// TIA Portal V20 export
// export: Created 2026-10-12T05:35:25.4874233Z, ExportSetting WithDefaults, DisplayName Totally Integrated Automation Portal, DisplayVersion V20, DisplayName TIA Portal Openness, DisplayVersion V20, DisplayName TIA Portal Teamcenter Gateway, DisplayVersion V20, DisplayName TIA Portal Version Control Interface, DisplayVersion V20, DisplayName SINAMICS Startdrive Advanced, DisplayVersion V20 SP1 Update 2, DisplayName SINAMICS Startdrive G110M, G120, G120C, G120D, G120P, G115D, DisplayVersion V20 SP1 Update 2, DisplayName SINAMICS Startdrive G130, G150, S120, S150, SINAMICS MV, G220, S200, S210, DisplayVersion V20 SP1 Update 2, DisplayName STEP 7 Professional, DisplayVersion V20, DisplayName STEP 7 Safety, DisplayVersion V20, DisplayName WinCC Basic/Comfort/Advanced, DisplayVersion V20, DisplayName WinCC Professional, DisplayVersion V20, DisplayName WinCC Unified, DisplayVersion V20
FUNCTION "FRK_ConfigFind" : Int   // FC96, SCL
{ S7_Optimized_Access := 'TRUE' }
VERSION : 0.1
// stored: AutoNumber true, IsIECCheckEnabled false, SetENOAutomatically false, UDAEnableTagReadback false
   VAR_INPUT
      Scope : String;
      Key : String;
      ModelCode : String;
   END_VAR
   VAR_TEMP
      Index : Int;
   END_VAR
BEGIN

   #FRK_ConfigFind := 0;
   FOR #Index := 1 TO 114 DO
       IF "FRK_ConfigStore".Rows[#Index].Used
           AND "FRK_ConfigStore".Rows[#Index].Record.Scope = #Scope
           AND "FRK_ConfigStore".Rows[#Index].Record.WriteKey = #Key
           AND "FRK_ConfigStore".Rows[#Index].ModelCode = #ModelCode THEN
           #FRK_ConfigFind := #Index;
           RETURN;
       END_IF;
   END_FOR;
END_FUNCTION
